Fanuc KAREL source: KA00107.KL

PROGRAM KA00107
%NOLOCKGROUP
VAR
  SRC: VECTOR
  DST: ARRAY[2] OF BYTE
BEGIN
  SRC.X = 1.0
  DST[1] = SRC
END KA00107
